TYPE stShutterCommand :
STRUCT
    CommandType  : eShutterCommandType;	// Command type
    Position : stShutterPosition;
END_STRUCT
END_TYPE

(* stored: Version 1.1.0.1
   DUT stShutterCommand: Id {23984a6c-c09a-4012-8087-64a064ebe57b} *)
